(*
SPDX-FileCopyrightText: © 2026 Oleksandr Tiutyk <trofimich@gmail.com>
SPDX-License-Identifier: MIT
License: https://opensource.org/license/mit
*)

(*!
<summary>Identifies an opaque configuration node within an active document.</summary>
<description>
Represents a node in a format-neutral hierarchical data model (JSON/YAML-style objects with named fields,
ordered arrays, or elementary values). Handles borrow the active document and expire when it is replaced or
closed. Do not store outside one synchronous load. Handle = 0 denotes an absent or unassigned node. Serialized
objects must ensure field names are unique within each object, safe for XML-like formats, and must not depend
on key order or case sensitivity.
</description>
*)
TYPE CONFIGURATION_NODE :
STRUCT
	Handle : __XWORD;
END_STRUCT
END_TYPE

(* stored: Version 1.1.0.1
   DUT CONFIGURATION_NODE: Id {c3b06388-c8df-485e-8350-b243242c1746} *)
